(* IEC 61131-3 sources: sis-interlock-demo/src/POUs/Sis/FB_SisEventLog, 5 files *)

(* ---- FB_SisEventLog.decl.st ---- *)
// Назначение: кольцевой журнал событий ПАЗ на SIS_LOG_SIZE записей: номер события udiSeq
//             присваивает журнал (1, 2, ...; после 16#FFFFFFFF — снова 1), самая старая запись
//             затирается. SCADA читает кольцо astRing по udiSeq и видит пропуски, если опрос
//             медленнее заполнения. Астрономическое время в ПЛК не ставится — дело приёмника.
// Автор:      kr0nsch
// Версия:     0.1.0
// Документ:   docs/DESIGN.md, раздел «7.1 FB_SisEventLog IMPLEMENTS I_SisEventSink»
// ВНИМАНИЕ:   код демонстрационный и не предназначен для систем безопасности. Реальная ПАЗ
//             требует определения SIL, сертифицированных аппаратных и программных средств
//             и валидации по ГОСТ Р МЭК 61511.
FUNCTION_BLOCK FB_SisEventLog IMPLEMENTS I_SisEventSink
VAR
    astRing : ARRAY[0..GVL_Const.SIS_LOG_SIZE - 1] OF ST_SisEvent;   // кольцо
    uiNext  : UINT;      // индекс следующей записи
    uiUsed  : UINT;      // занято, 0..SIS_LOG_SIZE
    udiSeq  : UDINT;     // номер последнего события
END_VAR

(* ---- AddEvent.method.decl.st ---- *)
// Записать событие с очередным номером (I_SisEventSink). Всегда TRUE: при заполнении кольца
// затирается самая старая запись
METHOD AddEvent : BOOL
VAR_INPUT
    stEvent : ST_SisEvent;   // событие; udiSeq заполняет журнал
END_VAR
VAR
    stRec : ST_SisEvent;     // запись с номером
END_VAR

(* ---- AddEvent.method.impl.st ---- *)
IF udiSeq = GVL_Const.UDINT_MAX THEN
    udiSeq := 1;
ELSE
    udiSeq := udiSeq + 1;
END_IF
stRec := stEvent;
stRec.udiSeq := udiSeq;
astRing[uiNext] := stRec;
uiNext := (uiNext + 1) MOD GVL_Const.SIS_LOG_SIZE;
IF uiUsed < GVL_Const.SIS_LOG_SIZE THEN
    uiUsed := uiUsed + 1;
END_IF
AddEvent := TRUE;

(* ---- GetEvent.method.decl.st ---- *)
// Событие uiBack записей назад (0 — последнее); uiBack >= Count — пустая запись (все поля 0)
METHOD GetEvent : ST_SisEvent
VAR_INPUT
    uiBack : UINT;           // сколько записей назад
END_VAR
VAR
    stEmpty : ST_SisEvent;   // пустая запись
    uiIdx   : UINT;          // индекс в кольце
END_VAR

(* ---- GetEvent.method.impl.st ---- *)
IF uiBack < uiUsed THEN
    // uiBack < uiUsed <= SIS_LOG_SIZE: выражение не уходит в минус
    uiIdx := (uiNext + GVL_Const.SIS_LOG_SIZE - 1 - uiBack) MOD GVL_Const.SIS_LOG_SIZE;
    GetEvent := astRing[uiIdx];
ELSE
    GetEvent := stEmpty;
END_IF
